FUNCTION_BLOCK ButtonM_HMI (* Service Interface Function Block Type *)
  (* Standard: 61499-2 *)
  (* Version 0.0, 6/20/2016, Andrei, nxtControl GmbH, template *)
  PACKAGE Main;
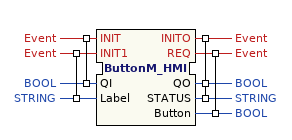
  EVENT_INPUT
    INIT WITH QI;
    INIT1 WITH Label;
  END_EVENT
  EVENT_OUTPUT
    INITO WITH QO, STATUS;
    REQ WITH Button;
  END_EVENT
  VAR_INPUT
    QI : BOOL;
    Label : STRING;
  END_VAR
  VAR_OUTPUT
    QO : BOOL; (* Event Output Qualifier *)
    STATUS : STRING; (* Service Status *)
    Button : BOOL;
  END_VAR
  SERVICE /
    SEQUENCE 
    END_SEQUENCE
  END_SERVICE
END_FUNCTION_BLOCK
